FUNCTION_BLOCK FB_DomeHomingState EXTENDS  FB_DomeState
VAR
END_VAR


METHOD CloseCommand : BOOL
// #202: a close is accepted in every state, it is the way to shut the roof
pDome^.SetState(pDome^.fbDomeCloseingState);
END_METHOD


PROPERTY StateID : STRING
GET
StateID := 'Homing State';
END_GET
END_PROPERTY

END_FUNCTION_BLOCK

(* stored: Version 1.1.0.1, ProductVersion 3.1.4024.15
   POU FB_DomeHomingState: Id {0b46cf97-8cde-4d7b-9e21-a3cae61e4b6e}, SpecialFunc None
   Method CloseCommand: Id {96eb34ec-9bda-4062-8e6e-6efc1b49e119}
   Property StateID: Id {ea9d5ebe-24bb-49b3-9665-3a8e0bb9c382}
   Get Get: Id {0414bc37-926c-4615-961d-e31436f44336} *)
